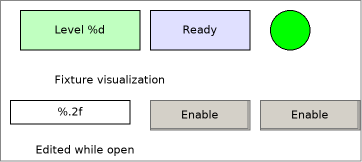
VISUALIZATION VISU_AllTypes  // 362x162
VAR_IN_OUT
	nLevel : INT;
	bFlag : BOOL;
END_VAR
    Rectangle (20,10 120x40), "Level %d", text variable: nLevel, colour toggle: GVL_Fixture.bEnable, invisible if: GVL_Fixture.bEnable, input disabled if: NOT GVL_Fixture.bEnable
        p3560616238: GVL_Fixture.nCount
        p2738717112: nLevel
        p2858320360: GVL_Fixture.nCount
    RoundedRectangle (150,10 100x40), "Ready"
    Ellipse (270,10 40x40), invisible if: GVL_Fixture.bEnable
    Label (10,70 200x20), "Fixture visualization"
    Textfield (10,100 120x24), "%.2f", text variable: GVL_Fixture.fValue
    Button (150,100 100x30), "Enable", tooltip "sets bEnable while pressed", pressed state: GVL_Fixture.bEnable
    Label (10,140 150x20), "Edited while open"
    Button (260,100 100x30), "Enable", tooltip "sets bEnable while pressed", pressed state: GVL_Fixture.bEnable
END_VISUALIZATION

(* stored: Version 1.1.0.1
   Visu VISU_AllTypes: Id {be1bb4c2-24e4-4d14-8a60-086936f9a6b7} *)
